// TIA Portal V20 export
// export: Created 2026-10-12T05:00:29.9809392Z, ExportSetting WithDefaults, DisplayName Totally Integrated Automation Portal, DisplayVersion V20, DisplayName TIA Portal Openness, DisplayVersion V20, DisplayName TIA Portal Teamcenter Gateway, DisplayVersion V20, DisplayName TIA Portal Version Control Interface, DisplayVersion V20, DisplayName SINAMICS Startdrive Advanced, DisplayVersion V20 SP1 Update 2, DisplayName SINAMICS Startdrive G110M, G120, G120C, G120D, G120P, G115D, DisplayVersion V20 SP1 Update 2, DisplayName SINAMICS Startdrive G130, G150, S120, S150, SINAMICS MV, G220, S200, S210, DisplayVersion V20 SP1 Update 2, DisplayName STEP 7 Professional, DisplayVersion V20, DisplayName STEP 7 Safety, DisplayVersion V20, DisplayName WinCC Basic/Comfort/Advanced, DisplayVersion V20, DisplayName WinCC Professional, DisplayVersion V20, DisplayName WinCC Unified, DisplayVersion V20
FUNCTION "FRK_SetFind" : Int   // FC105, SCL
{ S7_Optimized_Access := 'TRUE' }
VERSION : 0.1
// Deployment-sized keyed set storage; validation belongs to the typed walk.
// stored: AutoNumber true, IsIECCheckEnabled false, SetENOAutomatically false, UDAEnableTagReadback false
   VAR_INPUT
      RootIndex : Int;
      SetName : String;
   END_VAR
   VAR_TEMP
      Index : Int;
   END_VAR
BEGIN

   #FRK_SetFind := 0;
   FOR #Index := 1 TO 4 DO
       IF "FRK_SetStore".Sets[#RootIndex, #Index].Info.Used AND "FRK_SetStore".Sets[#RootIndex, #Index].Info.SetName = #SetName THEN
           #FRK_SetFind := #Index;
           RETURN;
       END_IF;
   END_FOR;
END_FUNCTION
